Staubli VAL3: goHome.pgx

public program goHome()
begin
  //stopMove()
  if !isEmpty()
    resetMotion()
  endIf
  movej(herej(),flange,mSimulate)
  movej(savedata:jHome,flange,mSimulate)
  waitEndMove()
end
